(* IEC 61131-3 sources: rusty/tests/lit/multi/polymorphism_interface, 7 files *)

(* ---- ia.st ---- *)
INTERFACE IA
    METHOD describeA : DINT
    END_METHOD
END_INTERFACE

(* ---- ib.st ---- *)
INTERFACE IB
    METHOD describeB : DINT
    END_METHOD
END_INTERFACE

(* ---- ic.st ---- *)
INTERFACE IC
    METHOD describeC : DINT
    END_METHOD
END_INTERFACE

(* ---- main.st ---- *)
FUNCTION main
    VAR
        instA: FbA;
        instB: FbB;
        instC: FbC;

        arrA: ARRAY[1..3] OF IA;
        arrB: ARRAY[1..2] OF IB;
        arrC: ARRAY[1..1] OF IC;

        i: DINT;
    END_VAR

    // All three FBs implement IA
    arrA[1] := instA;
    arrA[2] := instB;
    arrA[3] := instC;

    FOR i := 1 TO 3 DO
        printf('arrA[%d].describeA()=%d$N', i, arrA[i].describeA());
    END_FOR;

    // FbB and FbC implement IB
    arrB[1] := instB;
    arrB[2] := instC;

    FOR i := 1 TO 2 DO
        printf('arrB[%d].describeB()=%d$N', i, arrB[i].describeB());
    END_FOR;

    // Only FbC implements IC
    arrC[1] := instC;

    printf('arrC[1].describeC()=%d$N', arrC[1].describeC());
END_FUNCTION

(* ---- fb_a.st ---- *)
FUNCTION_BLOCK FbA IMPLEMENTS IA
    METHOD describeA : DINT
        printf('FbA::describeA$N');
        describeA := 1;
    END_METHOD
END_FUNCTION_BLOCK

(* ---- fb_b.st ---- *)
FUNCTION_BLOCK FbB IMPLEMENTS IA, IB
    METHOD describeA : DINT
        printf('FbB::describeA$N');
        describeA := 2;
    END_METHOD

    METHOD describeB : DINT
        printf('FbB::describeB$N');
        describeB := 20;
    END_METHOD
END_FUNCTION_BLOCK

(* ---- fb_c.st ---- *)
FUNCTION_BLOCK FbC IMPLEMENTS IA, IB, IC
    METHOD describeA : DINT
        printf('FbC::describeA$N');
        describeA := 3;
    END_METHOD

    METHOD describeB : DINT
        printf('FbC::describeB$N');
        describeB := 30;
    END_METHOD

    METHOD describeC : DINT
        printf('FbC::describeC$N');
        describeC := 300;
    END_METHOD
END_FUNCTION_BLOCK
